// TIA Portal V20 export
Screen "ProductionCount"  1276x673
  ScreenItem "Symbolic IO field_1" at 14,70 size 400x72  Type=HmiSymbolicIOField
  ScreenItem "Casella di testo_26" at 4,6 size 1273x53  Type=HmiTextBox
  ScreenItem "Casella di testo_14" at 864,147 size 400x34  Type=HmiTextBox
  ScreenItem "IO 域_82" at 864,217 size 106x34  Type=HmiIOField
  ScreenItem "IO 域_83" at 972,217 size 96x34  Type=HmiIOField
  ScreenItem "IO 域_84" at 1070,217 size 96x34  Type=HmiIOField
  ScreenItem "IO 域_85" at 1168,217 size 96x34  Type=HmiIOField
  ScreenItem "Casella di testo_21" at 864,183 size 106x34  Type=HmiTextBox
  ScreenItem "Casella di testo_23" at 972,183 size 96x34  Type=HmiTextBox
  ScreenItem "Casella di testo_24" at 1070,183 size 96x34  Type=HmiTextBox
  ScreenItem "Casella di testo_25" at 1168,183 size 96x34  Type=HmiTextBox
  ScreenItem "IO 域_86" at 864,252 size 106x34  Type=HmiIOField
  ScreenItem "IO 域_87" at 972,252 size 96x34  Type=HmiIOField
  ScreenItem "IO 域_88" at 1070,252 size 96x34  Type=HmiIOField
  ScreenItem "IO 域_89" at 1168,252 size 96x34  Type=HmiIOField
  ScreenItem "IO 域_90" at 864,287 size 106x34  Type=HmiIOField
  ScreenItem "IO 域_92" at 972,287 size 96x34  Type=HmiIOField
  ScreenItem "IO 域_93" at 1070,287 size 96x34  Type=HmiIOField
  ScreenItem "IO 域_94" at 1168,287 size 96x34  Type=HmiIOField
  ScreenItem "IO 域_95" at 864,323 size 106x34  Type=HmiIOField
  ScreenItem "IO 域_96" at 972,323 size 96x34  Type=HmiIOField
  ScreenItem "IO 域_97" at 1070,323 size 96x34  Type=HmiIOField
  ScreenItem "IO 域_98" at 1168,323 size 96x34  Type=HmiIOField
  ScreenItem "IO 域_120" at 864,359 size 106x34  Type=HmiIOField
  ScreenItem "IO 域_122" at 972,359 size 96x34  Type=HmiIOField
  ScreenItem "IO 域_123" at 1070,359 size 96x34  Type=HmiIOField
  ScreenItem "IO 域_81" at 1168,359 size 96x34  Type=HmiIOField
  ScreenItem "IO 域_124" at 864,394 size 106x34  Type=HmiIOField
  ScreenItem "IO 域_80" at 972,394 size 96x34  Type=HmiIOField
  ScreenItem "IO 域_78" at 1070,394 size 96x34  Type=HmiIOField
  ScreenItem "IO 域_45" at 1168,394 size 96x34  Type=HmiIOField
  ScreenItem "IO 域_46" at 864,429 size 106x34  Type=HmiIOField
  ScreenItem "IO 域_47" at 972,429 size 96x34  Type=HmiIOField
  ScreenItem "IO 域_48" at 1070,429 size 96x34  Type=HmiIOField
  ScreenItem "IO 域_49" at 1168,429 size 96x34  Type=HmiIOField
  ScreenItem "IO 域_51" at 864,464 size 106x34  Type=HmiIOField
  ScreenItem "IO 域_52" at 972,464 size 96x34  Type=HmiIOField
  ScreenItem "IO 域_53" at 1070,464 size 96x34  Type=HmiIOField
  ScreenItem "IO 域_54" at 1168,464 size 96x34  Type=HmiIOField
  ScreenItem "IO 域_66" at 864,552 size 132x46  Type=HmiIOField
  ScreenItem "Casella di testo_15" at 864,535 size 132x17  Type=HmiTextBox
  ScreenItem "IO 域_68" at 998,552 size 132x46  Type=HmiIOField
  ScreenItem "Casella di testo_17" at 998,535 size 132x17  Type=HmiTextBox
  ScreenItem "IO 域_69" at 998,621 size 132x46  Type=HmiIOField
  ScreenItem "Casella di testo_18" at 998,602 size 132x17  Type=HmiTextBox
  ScreenItem "IO 域_71" at 864,621 size 132x46  Type=HmiIOField
  ScreenItem "Casella di testo_19" at 864,602 size 132x17  Type=HmiTextBox
  ScreenItem "IO 域_72" at 1131,621 size 132x46  Type=HmiIOField
  ScreenItem "Casella di testo_20" at 1131,602 size 132x17  Type=HmiTextBox
  ScreenItem "IO 域_79" at 1131,552 size 132x46  Type=HmiIOField
  ScreenItem "Casella di testo_29" at 1131,535 size 132x17  Type=HmiTextBox
  ScreenItem "Casella di testo_1" at 438,147 size 400x34  Type=HmiTextBox
  ScreenItem "IO 域_25" at 438,217 size 106x34  Type=HmiIOField
  ScreenItem "IO 域_26" at 546,217 size 96x34  Type=HmiIOField
  ScreenItem "IO 域_27" at 644,217 size 96x34  Type=HmiIOField
  ScreenItem "IO 域_28" at 742,217 size 96x34  Type=HmiIOField
  ScreenItem "Casella di testo_8" at 438,183 size 106x34  Type=HmiTextBox
  ScreenItem "Casella di testo_9" at 546,183 size 96x34  Type=HmiTextBox
  ScreenItem "Casella di testo_10" at 644,183 size 96x34  Type=HmiTextBox
  ScreenItem "Casella di testo_12" at 742,183 size 96x34  Type=HmiTextBox
  ScreenItem "IO 域_29" at 438,252 size 106x34  Type=HmiIOField
  ScreenItem "IO 域_30" at 546,252 size 96x34  Type=HmiIOField
  ScreenItem "IO 域_31" at 644,252 size 96x34  Type=HmiIOField
  ScreenItem "IO 域_32" at 742,252 size 96x34  Type=HmiIOField
  ScreenItem "IO 域_33" at 438,287 size 106x34  Type=HmiIOField
  ScreenItem "IO 域_34" at 546,287 size 96x34  Type=HmiIOField
  ScreenItem "IO 域_35" at 644,287 size 96x34  Type=HmiIOField
  ScreenItem "IO 域_36" at 742,287 size 96x34  Type=HmiIOField
  ScreenItem "IO 域_37" at 438,323 size 106x34  Type=HmiIOField
  ScreenItem "IO 域_38" at 546,323 size 96x34  Type=HmiIOField
  ScreenItem "IO 域_39" at 644,323 size 96x34  Type=HmiIOField
  ScreenItem "IO 域_40" at 742,323 size 96x34  Type=HmiIOField
  ScreenItem "IO 域_41" at 438,359 size 106x34  Type=HmiIOField
  ScreenItem "IO 域_42" at 546,359 size 96x34  Type=HmiIOField
  ScreenItem "IO 域_43" at 644,359 size 96x34  Type=HmiIOField
  ScreenItem "IO 域_24" at 742,359 size 96x34  Type=HmiIOField
  ScreenItem "IO 域_44" at 438,394 size 106x34  Type=HmiIOField
  ScreenItem "IO 域_23" at 546,394 size 96x34  Type=HmiIOField
  ScreenItem "IO 域_21" at 644,394 size 96x34  Type=HmiIOField
  ScreenItem "IO 域_2" at 742,394 size 96x34  Type=HmiIOField
  ScreenItem "IO 域_4" at 438,429 size 106x34  Type=HmiIOField
  ScreenItem "IO 域_5" at 546,429 size 96x34  Type=HmiIOField
  ScreenItem "IO 域_6" at 644,429 size 96x34  Type=HmiIOField
  ScreenItem "IO 域_7" at 742,429 size 96x34  Type=HmiIOField
  ScreenItem "IO 域_8" at 438,464 size 106x34  Type=HmiIOField
  ScreenItem "IO 域_9" at 546,464 size 96x34  Type=HmiIOField
  ScreenItem "IO 域_10" at 644,464 size 96x34  Type=HmiIOField
  ScreenItem "IO 域_11" at 742,464 size 96x34  Type=HmiIOField
  ScreenItem "IO 域_12" at 438,499 size 106x34  Type=HmiIOField
  ScreenItem "IO 域_13" at 546,499 size 96x34  Type=HmiIOField
  ScreenItem "IO 域_14" at 644,499 size 96x34  Type=HmiIOField
  ScreenItem "IO 域_15" at 742,499 size 96x34  Type=HmiIOField
  ScreenItem "IO 域_16" at 438,552 size 132x46  Type=HmiIOField
  ScreenItem "Casella di testo_2" at 438,535 size 132x17  Type=HmiTextBox
  ScreenItem "IO 域_17" at 572,552 size 132x46  Type=HmiIOField
  ScreenItem "Casella di testo_3" at 572,535 size 132x17  Type=HmiTextBox
  ScreenItem "IO 域_18" at 572,621 size 132x46  Type=HmiIOField
  ScreenItem "Casella di testo_4" at 572,602 size 132x17  Type=HmiTextBox
  ScreenItem "IO 域_19" at 438,621 size 132x46  Type=HmiIOField
  ScreenItem "Casella di testo_5" at 438,602 size 132x17  Type=HmiTextBox
  ScreenItem "IO 域_20" at 705,621 size 132x46  Type=HmiIOField
  ScreenItem "Casella di testo_6" at 705,602 size 132x17  Type=HmiTextBox
  ScreenItem "IO 域_22" at 705,552 size 132x46  Type=HmiIOField
  ScreenItem "Casella di testo_13" at 705,535 size 132x17  Type=HmiTextBox
  ScreenItem "Casella di testo_47" at 14,147 size 400x34  Type=HmiTextBox
  ScreenItem "IO 域_76" at 14,217 size 106x34  Type=HmiIOField
  ScreenItem "IO 域_77" at 122,217 size 96x34  Type=HmiIOField
  ScreenItem "IO 域_55" at 220,217 size 96x34  Type=HmiIOField
  ScreenItem "IO 域_56" at 318,217 size 96x34  Type=HmiIOField
  ScreenItem "Casella di testo_43" at 14,183 size 106x34  Type=HmiTextBox
  ScreenItem "Casella di testo_49" at 122,183 size 96x34  Type=HmiTextBox
  ScreenItem "Casella di testo_27" at 220,183 size 96x34  Type=HmiTextBox
  ScreenItem "Casella di testo_28" at 318,183 size 96x34  Type=HmiTextBox
  ScreenItem "IO 域_57" at 14,252 size 106x34  Type=HmiIOField
  ScreenItem "IO 域_60" at 122,252 size 96x34  Type=HmiIOField
  ScreenItem "IO 域_61" at 220,252 size 96x34  Type=HmiIOField
  ScreenItem "IO 域_62" at 318,252 size 96x34  Type=HmiIOField
  ScreenItem "IO 域_65" at 14,287 size 106x34  Type=HmiIOField
  ScreenItem "IO 域_67" at 122,287 size 96x34  Type=HmiIOField
  ScreenItem "IO 域_70" at 220,287 size 96x34  Type=HmiIOField
  ScreenItem "IO 域_73" at 318,287 size 96x34  Type=HmiIOField
  ScreenItem "IO 域_74" at 14,323 size 106x34  Type=HmiIOField
  ScreenItem "IO 域_75" at 122,323 size 96x34  Type=HmiIOField
  ScreenItem "IO 域_99" at 220,323 size 96x34  Type=HmiIOField
  ScreenItem "IO 域_100" at 318,323 size 96x34  Type=HmiIOField
  ScreenItem "IO 域_103" at 14,359 size 106x34  Type=HmiIOField
  ScreenItem "IO 域_104" at 122,359 size 96x34  Type=HmiIOField
  ScreenItem "IO 域_105" at 220,359 size 96x34  Type=HmiIOField
  ScreenItem "IO 域_106" at 318,359 size 96x34  Type=HmiIOField
  ScreenItem "IO 域_107" at 14,394 size 106x34  Type=HmiIOField
  ScreenItem "IO 域_108" at 122,394 size 96x34  Type=HmiIOField
  ScreenItem "IO 域_109" at 220,394 size 96x34  Type=HmiIOField
  ScreenItem "IO 域_110" at 318,394 size 96x34  Type=HmiIOField
  ScreenItem "IO 域_111" at 14,429 size 106x34  Type=HmiIOField
  ScreenItem "IO 域_112" at 122,429 size 96x34  Type=HmiIOField
  ScreenItem "IO 域_113" at 220,429 size 96x34  Type=HmiIOField
  ScreenItem "IO 域_114" at 318,429 size 96x34  Type=HmiIOField
  ScreenItem "IO 域_115" at 14,464 size 106x34  Type=HmiIOField
  ScreenItem "IO 域_116" at 122,464 size 96x34  Type=HmiIOField
  ScreenItem "IO 域_117" at 220,464 size 96x34  Type=HmiIOField
  ScreenItem "IO 域_118" at 318,464 size 96x34  Type=HmiIOField
  ScreenItem "IO 域_101" at 14,499 size 106x34  Type=HmiIOField
  ScreenItem "IO 域_102" at 122,499 size 96x34  Type=HmiIOField
  ScreenItem "IO 域_119" at 220,499 size 96x34  Type=HmiIOField
  ScreenItem "IO 域_121" at 318,499 size 96x34  Type=HmiIOField
  ScreenItem "IO 域_162" at 14,552 size 132x46  Type=HmiIOField
  ScreenItem "Casella di testo_69" at 14,535 size 132x17  Type=HmiTextBox
  ScreenItem "IO 域_171" at 148,552 size 132x46  Type=HmiIOField
  ScreenItem "Casella di testo_72" at 148,535 size 132x17  Type=HmiTextBox
  ScreenItem "IO 域_164" at 148,621 size 132x46  Type=HmiIOField
  ScreenItem "Casella di testo_70" at 148,602 size 132x17  Type=HmiTextBox
  ScreenItem "IO 域_3" at 14,621 size 132x46  Type=HmiIOField
  ScreenItem "Casella di testo_11" at 14,602 size 132x17  Type=HmiTextBox
  ScreenItem "IO 域_161" at 281,621 size 132x46  Type=HmiIOField
  ScreenItem "Casella di testo_68" at 281,602 size 132x17  Type=HmiTextBox
  ScreenItem "IO 域_50" at 281,552 size 132x46  Type=HmiIOField
  ScreenItem "Casella di testo_22" at 281,535 size 132x17  Type=HmiTextBox
  ScreenItem "IO 域_244" at 440,90 size 176x52  Type=HmiIOField
  ScreenItem "Casella di testo_55" at 440,70 size 176x19  Type=HmiTextBox
  ScreenItem "IO 域_243" at 620,90 size 176x52  Type=HmiIOField
  ScreenItem "Casella di testo_53" at 620,70 size 176x19  Type=HmiTextBox
  ScreenItem "IO 域_91" at 801,90 size 176x52  Type=HmiIOField
  ScreenItem "Casella di testo_16" at 801,70 size 176x19  Type=HmiTextBox
  ScreenItem "IO 域_1" at 983,89 size 176x52  Type=HmiIOField
  ScreenItem "Casella di testo_7" at 983,69 size 176x19  Type=HmiTextBox
  ScreenItem "Button_15" at 1161,69 size 102x72  Type=HmiButton
